// TIA Portal V21 export
ORGANIZATION_BLOCK "OB_Dosing"   // OB124, SCL, ProgramCycle
TITLE = "Main Program Sweep (Cycle)" / Dosing cycle
// Program cycle OB of the unit Dosing; calls FB_Doser
// stored: Namespace Dosing, SetENOAutomatically false
   VAR_INPUT
      Initial_Call : Bool;   // Initial call of this OB
      Remanence : Bool;   // =True, if remanent data are available
   END_VAR
BEGIN

       "Dosing.IDB_Doser"(Start := TRUE, Stop := FALSE);
END_ORGANIZATION_BLOCK
